Staubli VAL3: new.pgx

public program new(string x_sKey, num x_nFrameIndex, num x_nToolIndex, num x_nMoveID, bool& x_bToSave)
begin
  if !isDefined(trajTemp:tTrajItem[x_sKey]) and x_sKey!=""
    insert(trajTemp:tTrajItem[x_sKey])
    trajTemp:tTrajItem[x_sKey].nFrameIndex=x_nFrameIndex
    trajTemp:tTrajItem[x_sKey].nToolIndex=x_nToolIndex
    trajTemp:tTrajItem[x_sKey].nMoveID=x_nMoveID
    //trajTemp:libSave()
    x_bToSave=true
    delay(0)
  else
    userPageAlert("项目存在，请重新命名！")
  endIf
end
